Fanuc KAREL source: kb00023.KL

-- PROVISIONAL review KL for V770-1; original PC SHA256 3cbe44e644d5a471d9a586bc85cb6db66cfc43d624c5859c58e07e55be38a073
-- Incomplete behavior may be omitted. Consult companion uncertainty JSON. Do not deploy.
PROGRAM KB00023
%NOLOCKGROUP
BEGIN
  -- UNRESOLVED_PC offsets 5-12; opcodes 9D,23
  -- UNRESOLVED_PC offsets 17-24; opcodes 9D,23
  -- UNRESOLVED_PC offsets 29-45; opcodes 27,22,22,31
  -- UNRESOLVED_PC offsets 50-54; opcodes 7F
END KB00023
